(* Logix 5000 project; controller CIP vendor 1 type 14 code 106 rev 20.12; software revision 20.06; part 11 of 13 *)
(* tags used below, declared in another part *)
   Bit : BOOL[128];
   Level_Bits : BOOL[32];
   MOA_ON : DINT[10];
   OpCode_Pin : DINT[5];
   Panelview : INT[40];
   PID1 : PID;
   PID2 : PID;
   PID3 : PID;
   PID3_Timer : TIMER[4];
   PID_Button : DINT[5];
   PID_Button_ONS : DINT[5];
   PID_ONS : DINT[5];
   PID_Timer : TIMER[5];
   PV_Valve_Input_Status_IND : INT[10,16];
   Recipe : RECIPE[41];
   SCLD_Dryer_Duct_Temp : REAL;
   SCLD_Supply_Flow : REAL;
   SCLD_Supply_Temp : REAL;
   SP_Dryer_Temp : REAL;
   SP_Supply_Flow : REAL;
   SP_Supply_Temp : REAL;
   Utility_Button : DINT[5];
   Utility_Button_ONS : DINT[5];
   Utility_ONS : DINT[5];
   Utility_Out : DINT[5];
   Utility_Timer : TIMER[20];
(* MainProgram, continued *)

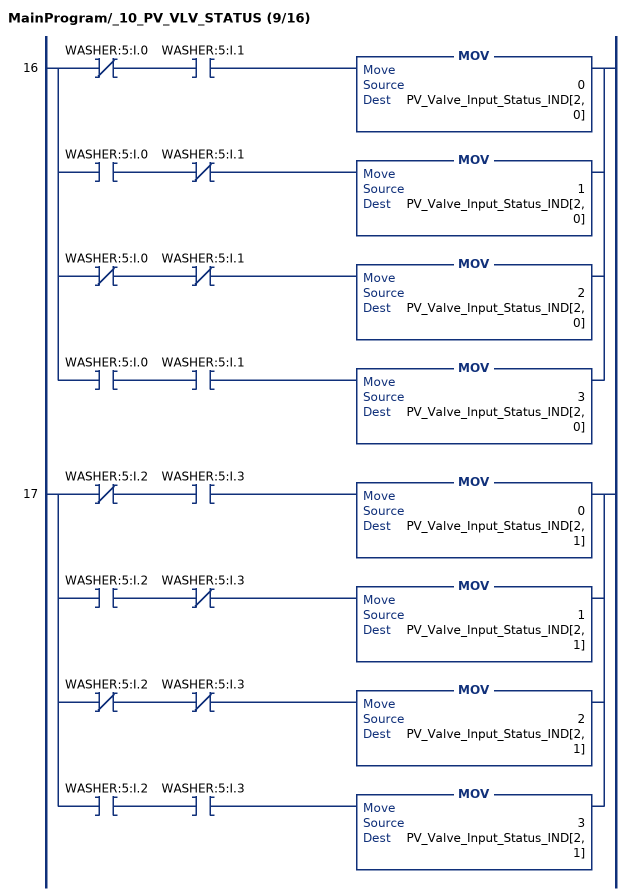
   [picture p205: MainProgram/_10_PV_VLV_STATUS rungs 16-17]
   16: [XIO(WASHER:5:I.0) XIC(WASHER:5:I.1) MOV(0,PV_Valve_Input_Status_IND[2,0]) ,XIC(WASHER:5:I.0) XIO(WASHER:5:I.1) MOV(1,PV_Valve_Input_Status_IND[2,0]) ,XIO(WASHER:5:I.0) XIO(WASHER:5:I.1) MOV(2,PV_Valve_Input_Status_IND[2,0]) ,XIC(WASHER:5:I.0) XIC(WASHER:5:I.1) MOV(3,PV_Valve_Input_Status_IND[2,0]) ];
   17: [XIO(WASHER:5:I.2) XIC(WASHER:5:I.3) MOV(0,PV_Valve_Input_Status_IND[2,1]) ,XIC(WASHER:5:I.2) XIO(WASHER:5:I.3) MOV(1,PV_Valve_Input_Status_IND[2,1]) ,XIO(WASHER:5:I.2) XIO(WASHER:5:I.3) MOV(2,PV_Valve_Input_Status_IND[2,1]) ,XIC(WASHER:5:I.2) XIC(WASHER:5:I.3) MOV(3,PV_Valve_Input_Status_IND[2,1]) ];
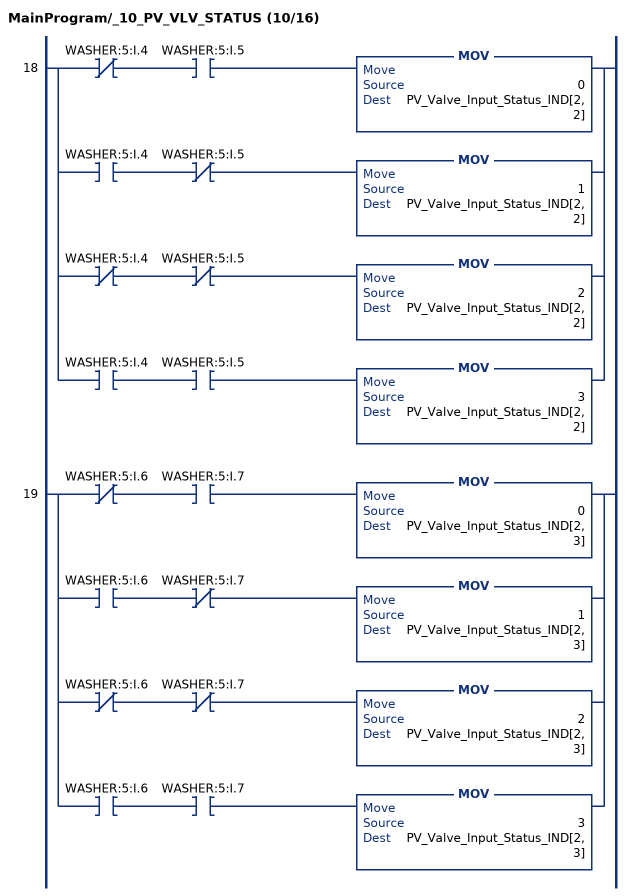
   18: [XIO(WASHER:5:I.4) XIC(WASHER:5:I.5) MOV(0,PV_Valve_Input_Status_IND[2,2]) ,XIC(WASHER:5:I.4) XIO(WASHER:5:I.5) MOV(1,PV_Valve_Input_Status_IND[2,2]) ,XIO(WASHER:5:I.4) XIO(WASHER:5:I.5) MOV(2,PV_Valve_Input_Status_IND[2,2]) ,XIC(WASHER:5:I.4) XIC(WASHER:5:I.5) MOV(3,PV_Valve_Input_Status_IND[2,2]) ];
   19: [XIO(WASHER:5:I.6) XIC(WASHER:5:I.7) MOV(0,PV_Valve_Input_Status_IND[2,3]) ,XIC(WASHER:5:I.6) XIO(WASHER:5:I.7) MOV(1,PV_Valve_Input_Status_IND[2,3]) ,XIO(WASHER:5:I.6) XIO(WASHER:5:I.7) MOV(2,PV_Valve_Input_Status_IND[2,3]) ,XIC(WASHER:5:I.6) XIC(WASHER:5:I.7) MOV(3,PV_Valve_Input_Status_IND[2,3]) ];
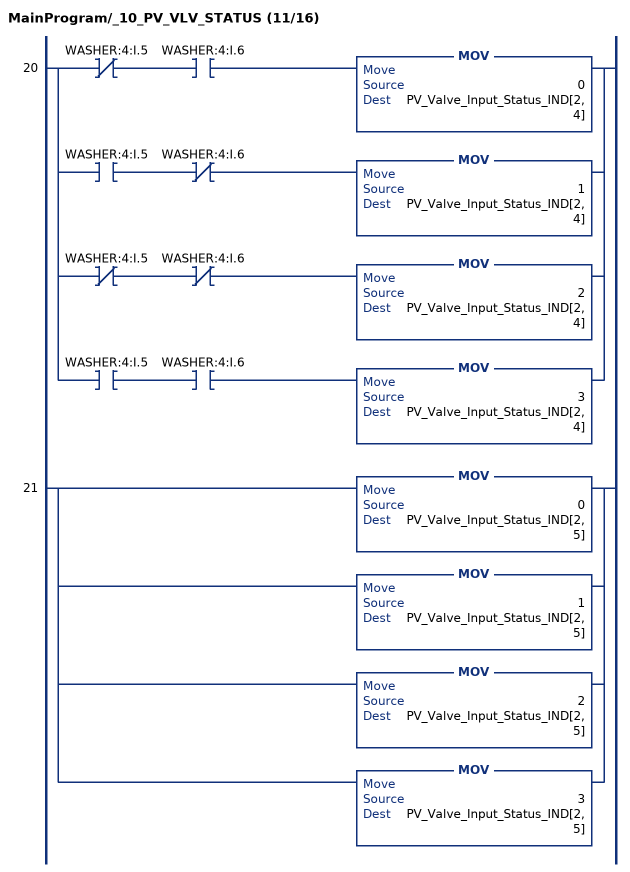
   20: [XIO(WASHER:4:I.5) XIC(WASHER:4:I.6) MOV(0,PV_Valve_Input_Status_IND[2,4]) ,XIC(WASHER:4:I.5) XIO(WASHER:4:I.6) MOV(1,PV_Valve_Input_Status_IND[2,4]) ,XIO(WASHER:4:I.5) XIO(WASHER:4:I.6) MOV(2,PV_Valve_Input_Status_IND[2,4]) ,XIC(WASHER:4:I.5) XIC(WASHER:4:I.6) MOV(3,PV_Valve_Input_Status_IND[2,4]) ];
   21: [MOV(0,PV_Valve_Input_Status_IND[2,5]) ,MOV(1,PV_Valve_Input_Status_IND[2,5]) ,MOV(2,PV_Valve_Input_Status_IND[2,5]) ,MOV(3,PV_Valve_Input_Status_IND[2,5]) ];
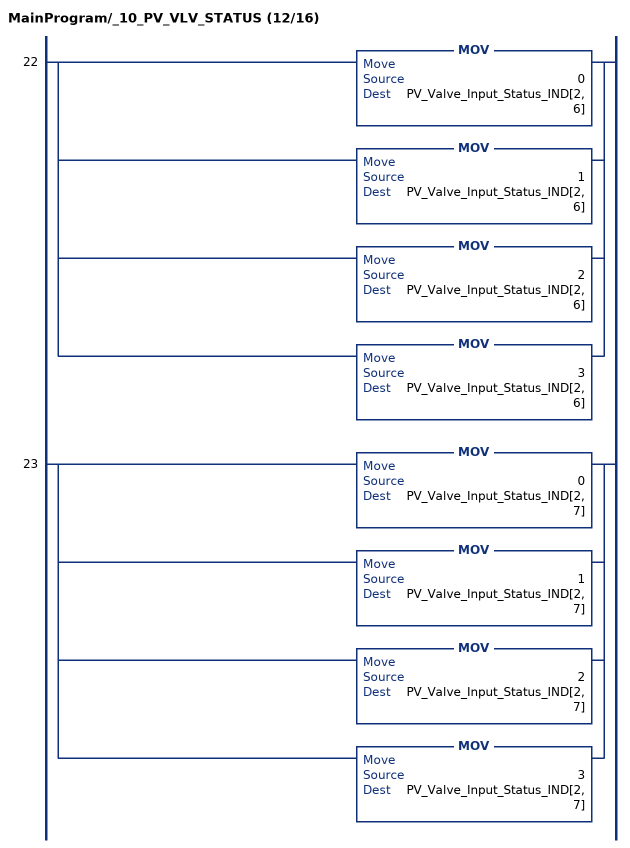
   22: [MOV(0,PV_Valve_Input_Status_IND[2,6]) ,MOV(1,PV_Valve_Input_Status_IND[2,6]) ,MOV(2,PV_Valve_Input_Status_IND[2,6]) ,MOV(3,PV_Valve_Input_Status_IND[2,6]) ];
   23: [MOV(0,PV_Valve_Input_Status_IND[2,7]) ,MOV(1,PV_Valve_Input_Status_IND[2,7]) ,MOV(2,PV_Valve_Input_Status_IND[2,7]) ,MOV(3,PV_Valve_Input_Status_IND[2,7]) ];
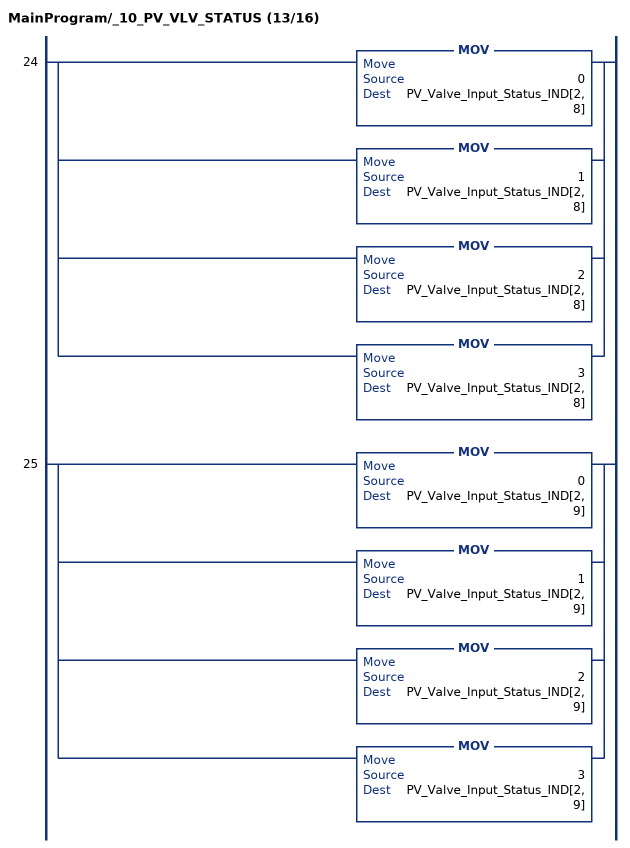
   24: [MOV(0,PV_Valve_Input_Status_IND[2,8]) ,MOV(1,PV_Valve_Input_Status_IND[2,8]) ,MOV(2,PV_Valve_Input_Status_IND[2,8]) ,MOV(3,PV_Valve_Input_Status_IND[2,8]) ];
   25: [MOV(0,PV_Valve_Input_Status_IND[2,9]) ,MOV(1,PV_Valve_Input_Status_IND[2,9]) ,MOV(2,PV_Valve_Input_Status_IND[2,9]) ,MOV(3,PV_Valve_Input_Status_IND[2,9]) ];
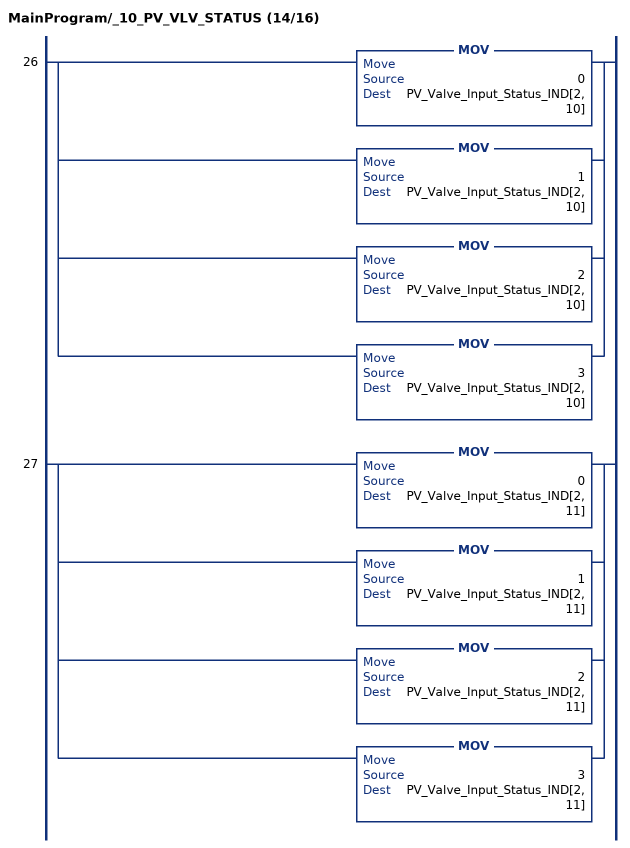
   26: [MOV(0,PV_Valve_Input_Status_IND[2,10]) ,MOV(1,PV_Valve_Input_Status_IND[2,10]) ,MOV(2,PV_Valve_Input_Status_IND[2,10]) ,MOV(3,PV_Valve_Input_Status_IND[2,10]) ];
   27: [MOV(0,PV_Valve_Input_Status_IND[2,11]) ,MOV(1,PV_Valve_Input_Status_IND[2,11]) ,MOV(2,PV_Valve_Input_Status_IND[2,11]) ,MOV(3,PV_Valve_Input_Status_IND[2,11]) ];
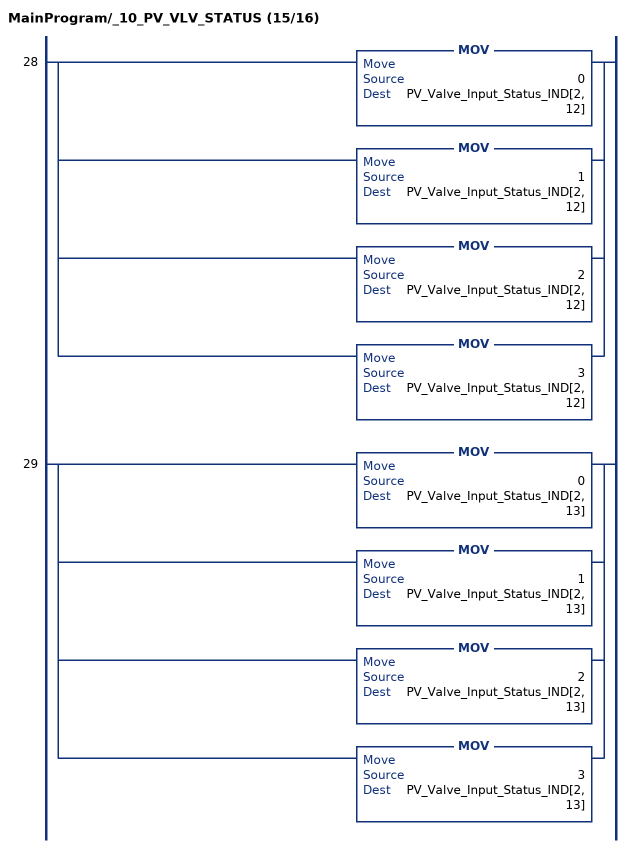
   28: [MOV(0,PV_Valve_Input_Status_IND[2,12]) ,MOV(1,PV_Valve_Input_Status_IND[2,12]) ,MOV(2,PV_Valve_Input_Status_IND[2,12]) ,MOV(3,PV_Valve_Input_Status_IND[2,12]) ];
   29: [MOV(0,PV_Valve_Input_Status_IND[2,13]) ,MOV(1,PV_Valve_Input_Status_IND[2,13]) ,MOV(2,PV_Valve_Input_Status_IND[2,13]) ,MOV(3,PV_Valve_Input_Status_IND[2,13]) ];
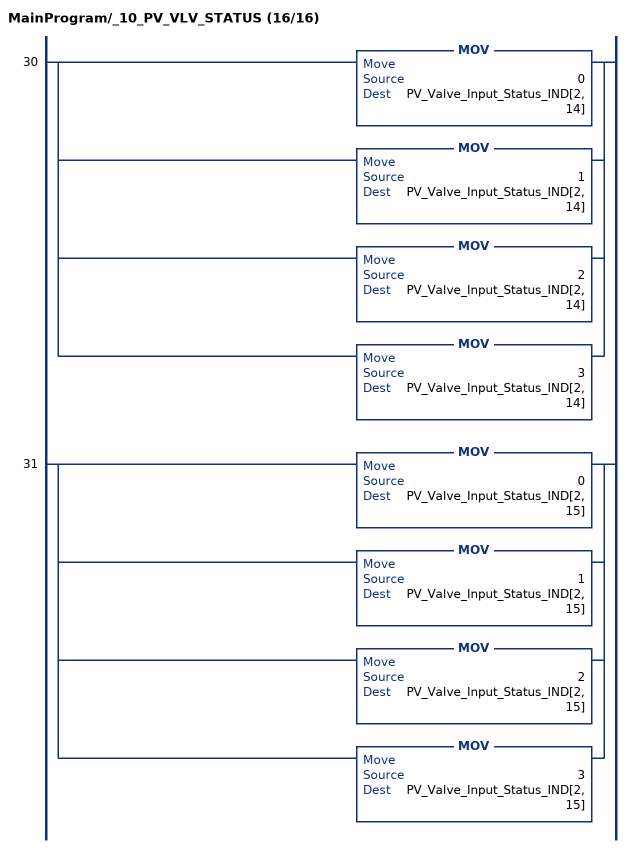
   30: [MOV(0,PV_Valve_Input_Status_IND[2,14]) ,MOV(1,PV_Valve_Input_Status_IND[2,14]) ,MOV(2,PV_Valve_Input_Status_IND[2,14]) ,MOV(3,PV_Valve_Input_Status_IND[2,14]) ];
   31: [MOV(0,PV_Valve_Input_Status_IND[2,15]) ,MOV(1,PV_Valve_Input_Status_IND[2,15]) ,MOV(2,PV_Valve_Input_Status_IND[2,15]) ,MOV(3,PV_Valve_Input_Status_IND[2,15]) ];
END_ROUTINE

ROUTINE _20_UTILITY   (* ladder *)
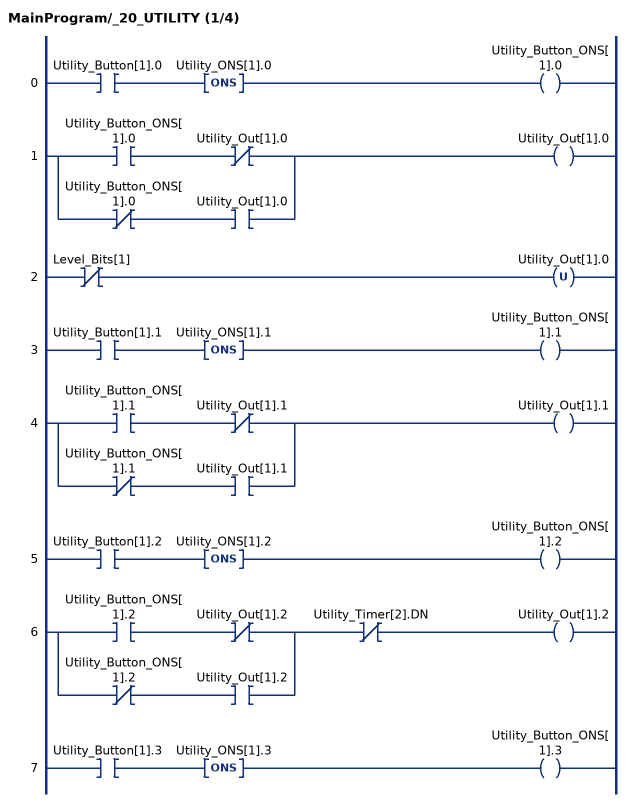
   0: XIC(Utility_Button[1].0)ONS(Utility_ONS[1].0)OTE(Utility_Button_ONS[1].0);
   1: [XIC(Utility_Button_ONS[1].0) XIO(Utility_Out[1].0) ,XIO(Utility_Button_ONS[1].0) XIC(Utility_Out[1].0) ]OTE(Utility_Out[1].0);
   2: XIO(Level_Bits[1])OTU(Utility_Out[1].0);
   3: XIC(Utility_Button[1].1)ONS(Utility_ONS[1].1)OTE(Utility_Button_ONS[1].1);
   4: [XIC(Utility_Button_ONS[1].1) XIO(Utility_Out[1].1) ,XIO(Utility_Button_ONS[1].1) XIC(Utility_Out[1].1) ]OTE(Utility_Out[1].1);
   5: XIC(Utility_Button[1].2)ONS(Utility_ONS[1].2)OTE(Utility_Button_ONS[1].2);
   6: [XIC(Utility_Button_ONS[1].2) XIO(Utility_Out[1].2) ,XIO(Utility_Button_ONS[1].2) XIC(Utility_Out[1].2) ]XIO(Utility_Timer[2].DN)OTE(Utility_Out[1].2);
   7: XIC(Utility_Button[1].3)ONS(Utility_ONS[1].3)OTE(Utility_Button_ONS[1].3);
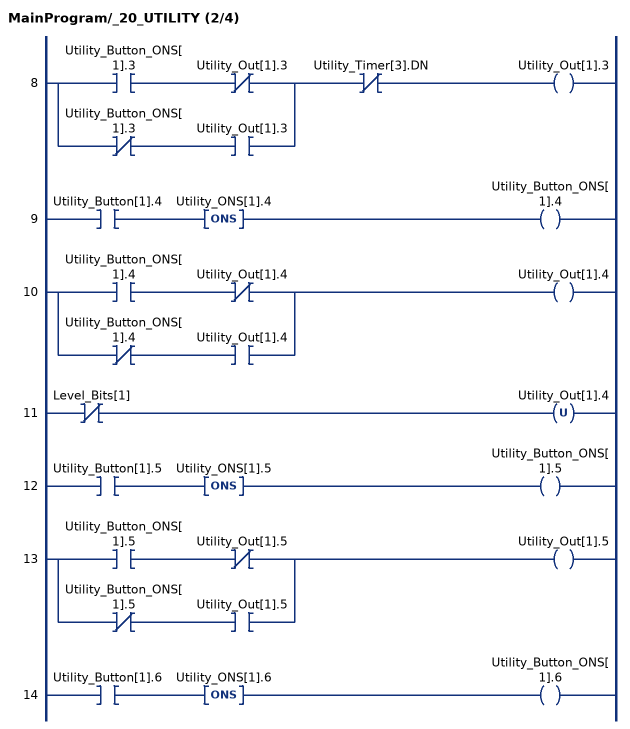
   8: [XIC(Utility_Button_ONS[1].3) XIO(Utility_Out[1].3) ,XIO(Utility_Button_ONS[1].3) XIC(Utility_Out[1].3) ]XIO(Utility_Timer[3].DN)OTE(Utility_Out[1].3);
   9: XIC(Utility_Button[1].4)ONS(Utility_ONS[1].4)OTE(Utility_Button_ONS[1].4);
   10: [XIC(Utility_Button_ONS[1].4) XIO(Utility_Out[1].4) ,XIO(Utility_Button_ONS[1].4) XIC(Utility_Out[1].4) ]OTE(Utility_Out[1].4);
   11: XIO(Level_Bits[1])OTU(Utility_Out[1].4);
   12: XIC(Utility_Button[1].5)ONS(Utility_ONS[1].5)OTE(Utility_Button_ONS[1].5);
   13: [XIC(Utility_Button_ONS[1].5) XIO(Utility_Out[1].5) ,XIO(Utility_Button_ONS[1].5) XIC(Utility_Out[1].5) ]OTE(Utility_Out[1].5);
   14: XIC(Utility_Button[1].6)ONS(Utility_ONS[1].6)OTE(Utility_Button_ONS[1].6);
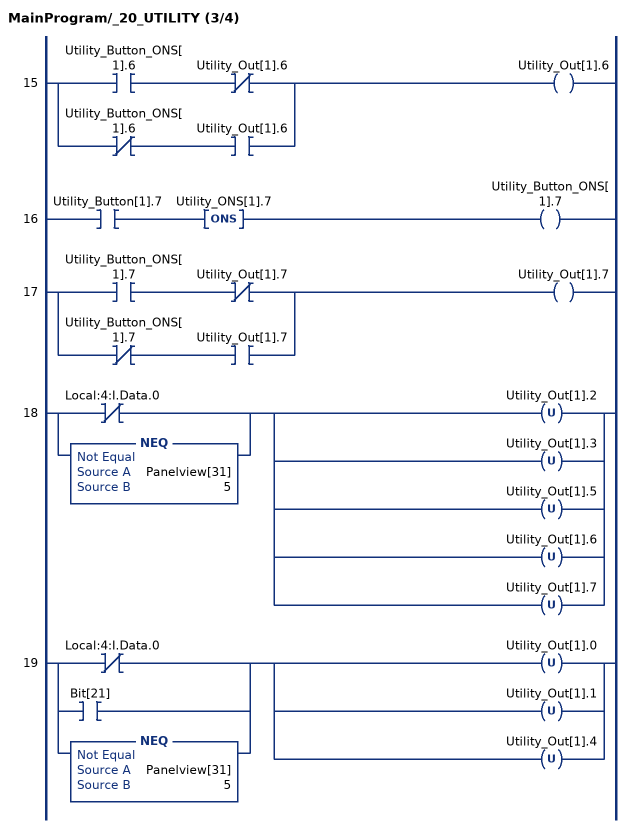
   15: [XIC(Utility_Button_ONS[1].6) XIO(Utility_Out[1].6) ,XIO(Utility_Button_ONS[1].6) XIC(Utility_Out[1].6) ]OTE(Utility_Out[1].6);
   16: XIC(Utility_Button[1].7)ONS(Utility_ONS[1].7)OTE(Utility_Button_ONS[1].7);
   17: [XIC(Utility_Button_ONS[1].7) XIO(Utility_Out[1].7) ,XIO(Utility_Button_ONS[1].7) XIC(Utility_Out[1].7) ]OTE(Utility_Out[1].7);
   18: [XIO(Local:4:I.Data.0) ,NEQ(Panelview[31],5) ][OTU(Utility_Out[1].2) ,OTU(Utility_Out[1].3) ,OTU(Utility_Out[1].5) ,OTU(Utility_Out[1].6) ,OTU(Utility_Out[1].7) ];
   19: [XIO(Local:4:I.Data.0) ,XIC(Bit[21]) ,NEQ(Panelview[31],5) ][OTU(Utility_Out[1].0) ,OTU(Utility_Out[1].1) ,OTU(Utility_Out[1].4) ];
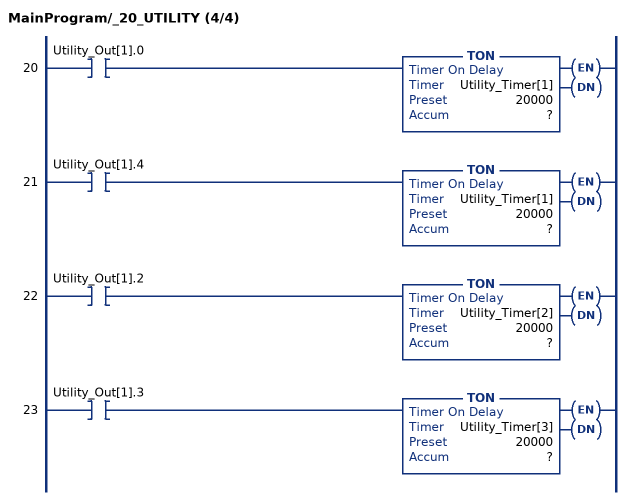
   20: XIC(Utility_Out[1].0)TON(Utility_Timer[1],?,?);
   21: XIC(Utility_Out[1].4)TON(Utility_Timer[1],?,?);
   22: XIC(Utility_Out[1].2)TON(Utility_Timer[2],?,?);
   23: XIC(Utility_Out[1].3)TON(Utility_Timer[3],?,?);
END_ROUTINE

ROUTINE _25_PID1_SUPPLY_TEMP   (* ladder *)
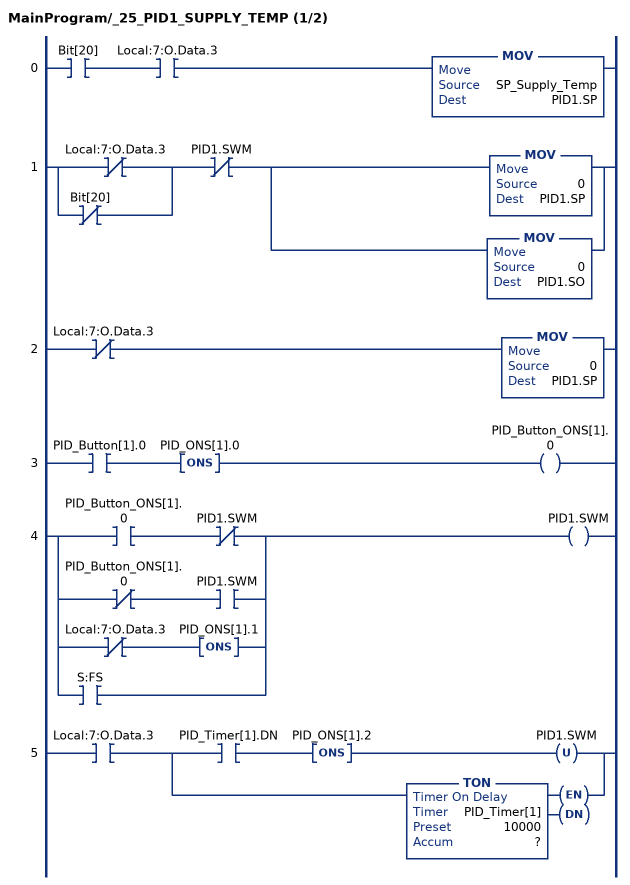
   0: XIC(Bit[20])XIC(Local:7:O.Data.3)MOV(SP_Supply_Temp,PID1.SP);
   1: [XIO(Local:7:O.Data.3) ,XIO(Bit[20]) ]XIO(PID1.SWM)[MOV(0,PID1.SP) ,MOV(0,PID1.SO) ];
   2: XIO(Local:7:O.Data.3)MOV(0,PID1.SP);
   3: XIC(PID_Button[1].0)ONS(PID_ONS[1].0)OTE(PID_Button_ONS[1].0);
   4: [XIC(PID_Button_ONS[1].0) XIO(PID1.SWM) ,XIO(PID_Button_ONS[1].0) XIC(PID1.SWM) ,XIO(Local:7:O.Data.3) ONS(PID_ONS[1].1) ,XIC(S:FS) ]OTE(PID1.SWM);
   5: XIC(Local:7:O.Data.3)[XIC(PID_Timer[1].DN) ONS(PID_ONS[1].2) OTU(PID1.SWM) ,TON(PID_Timer[1],?,?) ];
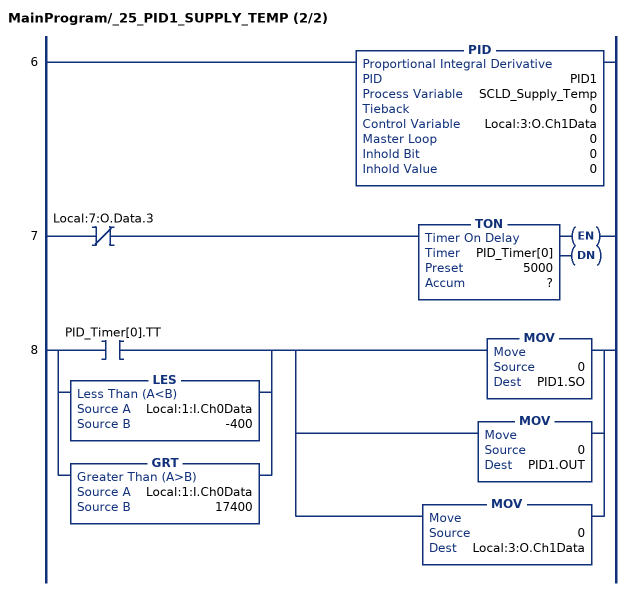
   6: PID(PID1,SCLD_Supply_Temp,0,Local:3:O.Ch1Data,0,0,0);
   7: XIO(Local:7:O.Data.3)TON(PID_Timer[0],?,?);
   8: [XIC(PID_Timer[0].TT) ,LES(Local:1:I.Ch0Data,-400) ,GRT(Local:1:I.Ch0Data,17400) ][MOV(0,PID1.SO) ,MOV(0,PID1.OUT) ,MOV(0,Local:3:O.Ch1Data) ];
END_ROUTINE

ROUTINE _25_PID2_SUPPLY_FLOW   (* ladder *)
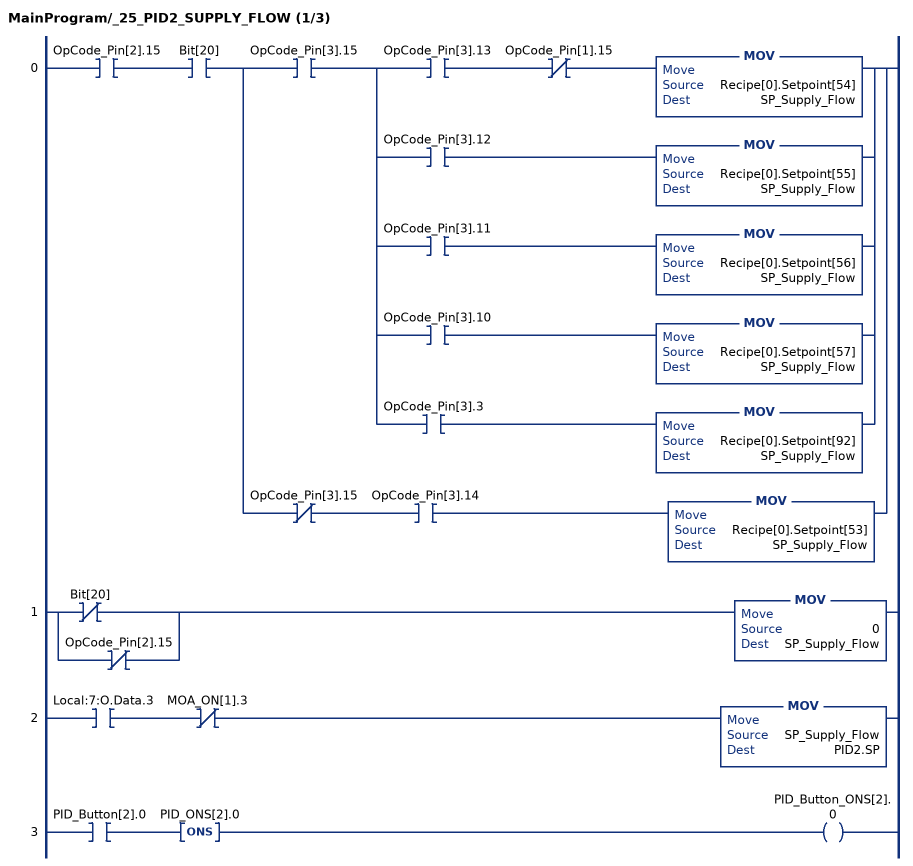
   0: XIC(OpCode_Pin[2].15)XIC(Bit[20])[XIC(OpCode_Pin[3].15) [XIC(OpCode_Pin[3].13) XIO(OpCode_Pin[1].15) MOV(Recipe[0].Setpoint[54],SP_Supply_Flow) ,XIC(OpCode_Pin[3].12) MOV(Recipe[0].Setpoint[55],SP_Supply_Flow) ,XIC(OpCode_Pin[3].11) MOV(Recipe[0].Setpoint[56],SP_Supply_Flow) ,XIC(OpCode_Pin[3].10) MOV(Recipe[0].Setpoint[57],SP_Supply_Flow) ,XIC(OpCode_Pin[3].3) MOV(Recipe[0].Setpoint[92],SP_Supply_Flow) ] ,XIO(OpCode_Pin[3].15) XIC(OpCode_Pin[3].14) MOV(Recipe[0].Setpoint[53],SP_Supply_Flow) ];
   1: [XIO(Bit[20]) ,XIO(OpCode_Pin[2].15) ]MOV(0,SP_Supply_Flow);
   2: XIC(Local:7:O.Data.3)XIO(MOA_ON[1].3)MOV(SP_Supply_Flow,PID2.SP);
   3: XIC(PID_Button[2].0)ONS(PID_ONS[2].0)OTE(PID_Button_ONS[2].0);
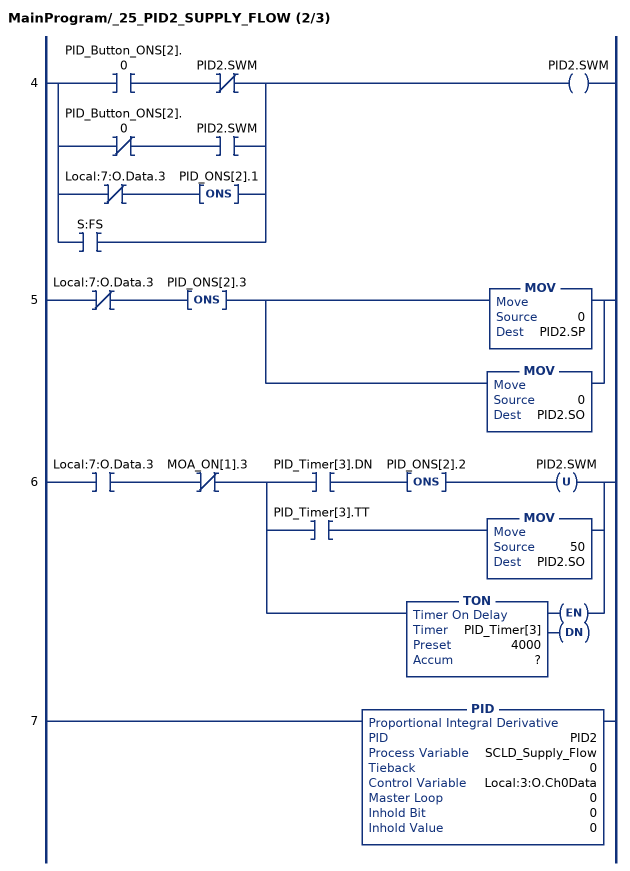
   4: [XIC(PID_Button_ONS[2].0) XIO(PID2.SWM) ,XIO(PID_Button_ONS[2].0) XIC(PID2.SWM) ,XIO(Local:7:O.Data.3) ONS(PID_ONS[2].1) ,XIC(S:FS) ]OTE(PID2.SWM);
   5: XIO(Local:7:O.Data.3)ONS(PID_ONS[2].3)[MOV(0,PID2.SP) ,MOV(0,PID2.SO) ];
   6: XIC(Local:7:O.Data.3)XIO(MOA_ON[1].3)[XIC(PID_Timer[3].DN) ONS(PID_ONS[2].2) OTU(PID2.SWM) ,XIC(PID_Timer[3].TT) MOV(50,PID2.SO) ,TON(PID_Timer[3],?,?) ];
   7: PID(PID2,SCLD_Supply_Flow,0,Local:3:O.Ch0Data,0,0,0);
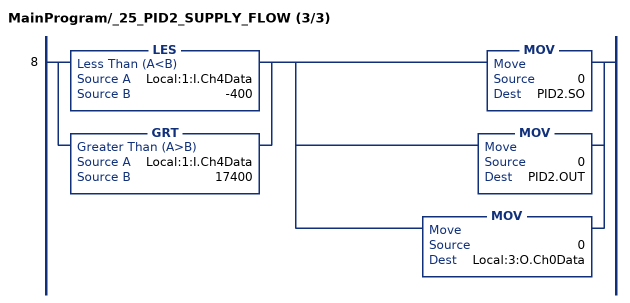
   8: [LES(Local:1:I.Ch4Data,-400) ,GRT(Local:1:I.Ch4Data,17400) ][MOV(0,PID2.SO) ,MOV(0,PID2.OUT) ,MOV(0,Local:3:O.Ch0Data) ];
END_ROUTINE

ROUTINE _25_PID3_DRYER_TEMP   (* ladder *)
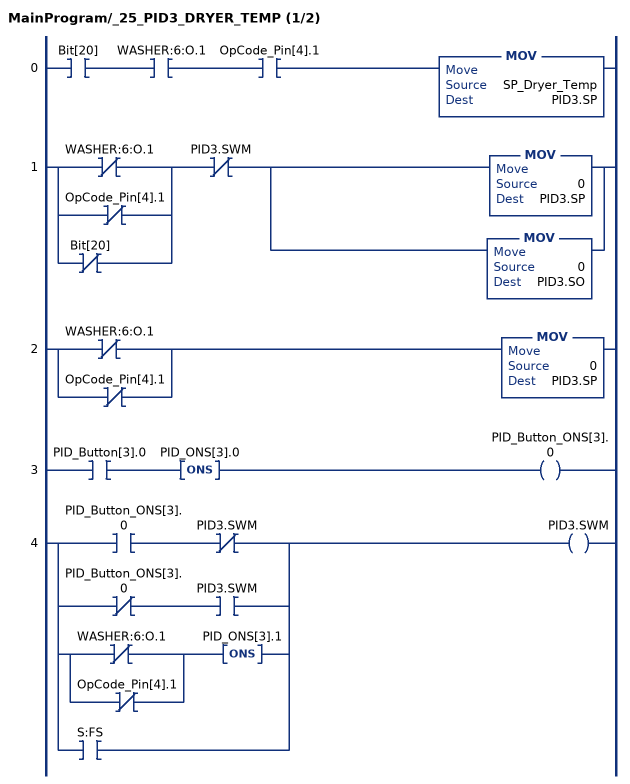
   0: XIC(Bit[20])XIC(WASHER:6:O.1)XIC(OpCode_Pin[4].1)MOV(SP_Dryer_Temp,PID3.SP);
   1: [XIO(WASHER:6:O.1) ,XIO(OpCode_Pin[4].1) ,XIO(Bit[20]) ]XIO(PID3.SWM)[MOV(0,PID3.SP) ,MOV(0,PID3.SO) ];
   2: [XIO(WASHER:6:O.1) ,XIO(OpCode_Pin[4].1) ]MOV(0,PID3.SP);
   3: XIC(PID_Button[3].0)ONS(PID_ONS[3].0)OTE(PID_Button_ONS[3].0);
   4: [XIC(PID_Button_ONS[3].0) XIO(PID3.SWM) ,XIO(PID_Button_ONS[3].0) XIC(PID3.SWM) ,[XIO(WASHER:6:O.1) ,XIO(OpCode_Pin[4].1) ] ONS(PID_ONS[3].1) ,XIC(S:FS) ]OTE(PID3.SWM);
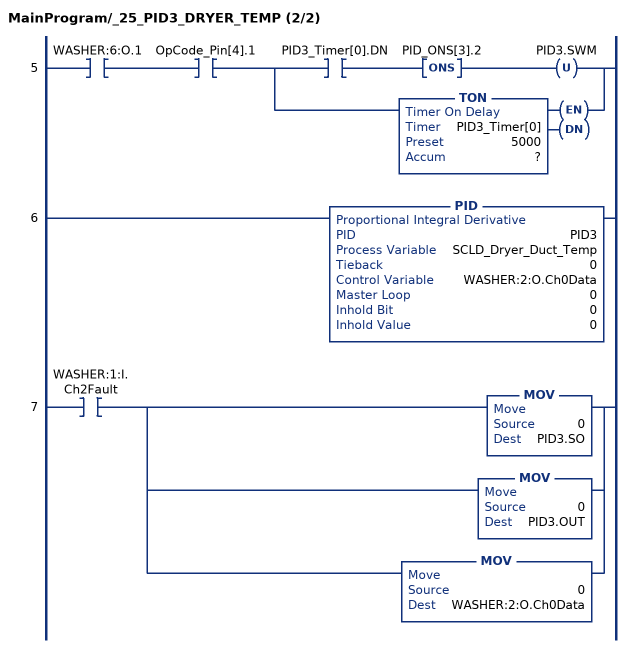
   5: XIC(WASHER:6:O.1)XIC(OpCode_Pin[4].1)[XIC(PID3_Timer[0].DN) ONS(PID_ONS[3].2) OTU(PID3.SWM) ,TON(PID3_Timer[0],?,?) ];
   6: PID(PID3,SCLD_Dryer_Duct_Temp,0,WASHER:2:O.Ch0Data,0,0,0);
   7: XIC(WASHER:1:I.Ch2Fault)[MOV(0,PID3.SO) ,MOV(0,PID3.OUT) ,MOV(0,WASHER:2:O.Ch0Data) ];
END_ROUTINE
